Staubli VAL3: refreshQuit.pgx

public program refreshQuit(bool& x_bOut)
begin
  //Quit
  if utBtn_Step[0].Events.bClick==false and  utBtn_Step[1].Events.bClick==false and utBtn_Step[2].Events.bClick==false and utBtn_Step[3].Events.bClick==false
    if utBtn_Bottom[7].Events.bClick==true
      utBtn_Bottom[7].Events.bClick=false
      //Press F7
      call hmiConfirm("Quit","confirm",x_bOut)
    endIf
  endIf
end
